Staubli VAL3: Matrix2Trsf.pgx

public program Matrix2Trsf(num& x_nMatrix[] (dimensions=2), trsf& x_trTrsf)
  local num ax
  local num ay
  local num az
  local num nx
  local num ny
  local num nz
  local num ox
  local num oy
  local num oz
  local num px
  local num py
  local num pz
  local num rx1
  local num rx2
  local num ry1
  local num ry2
  local num rz1
  local num rz2
  local num x
  local num y
  local num z
begin
  //Matrik转换成Trsf
  nx=x_nMatrix[0,0]
  ny=x_nMatrix[0,1]
  nz=x_nMatrix[0,2]
  ox=x_nMatrix[1,0]
  oy=x_nMatrix[1,1]
  oz=x_nMatrix[1,2]
  ax=x_nMatrix[2,0]
  ay=x_nMatrix[2,1]
  az=x_nMatrix[2,2]
  px=x_nMatrix[3,0]
  py=x_nMatrix[3,1]
  pz=x_nMatrix[3,2]
  //求解Rx、Ry、Rz
  x_trTrsf.x=px
  x_trTrsf.y=py
  x_trTrsf.z=pz
  //求解Rx、Ry、Rz
  call Atan2(ax,sqrt(power(nx,2)+power(ox,2)),ry1)
  if ry1==90
    rx1=0
    call Atan2(ny,-nz,rz1)
  elseIf ry1==-90
    rx1=0
    call Atan2(ny,nz,rz1)
  else
    call Atan2(-ay/cos(ry1),az/cos(ry1),rx1)
    call Atan2(-ox/cos(ry1),nx/cos(ry1),rz1)
  endIf

  call Atan2(ax,sqrt(power(nx,2)+power(ox,2)),ry2)
  if ry2==90
    rx2=0
    call Atan2(ny,-nz,rz2)
  elseIf ry2==-90
    rx2=0
    call Atan2(ny,nz,rz2)
  else
    call Atan2(-ay/cos(ry2),az/cos(ry2),rx2)
    call Atan2(-ox/cos(ry2),nx/cos(ry2),rz2)
  endIf

  if abs(rx1)+abs(ry1)+abs(rz1)<=abs(rx2)+abs(ry2)+abs(rz2)
    x_trTrsf.rx=rx1
    x_trTrsf.ry=ry1
    x_trTrsf.rz=rz1
  else
    x_trTrsf.rx=rx2
    x_trTrsf.ry=ry2
    x_trTrsf.rz=rz2
  endIf
end
